(* IEC 61131-3 sources: Elmo_Master/Lasal_PRG/Elmo_EtherCAT_Test_4Axis/Network, 1 file *)

(* ---- ConfigObjects.st ---- *)
FUNCTION GLOBAL TAB TASK_CONF
_K_TASK, _K_REAL,
_K_END_VAR,

_K_TASK, _K_CYCLIC,
_K_END_VAR,

_K_TASK, _K_BACKGROUND,
_K_END_VAR,

_K_END_CONF
END_FUNCTION

FUNCTION GLOBAL TAB IPR_CONF
_K_IPR
	0$UINT,
_K_END_VAR,
_K_END_CONF
END_FUNCTION

FUNCTION GLOBAL TAB CONFIG_TABLES
00121$UINT,
0$UINT, 1, 58, "_AXISBASE",
0$UINT, 0, 5, "_CAN",
0$UINT, 1, 11, "_CANLIB",
0$UINT, 1, 0, "_CHECKSUM",
0$UINT, 1, 20, "_FILESYS",
0$UINT, 0, 5, "_LINKER",
0$UINT, 1, 0, "_LMCABSENCODER",
0$UINT, 1, 120, "_LMCAXIS",
0$UINT, 2, 111, "_LMCAXISBASE",
0$UINT, 1, 32, "_LMCAXISREF",
0$UINT, 1, 42, "_LMCAXISVIS",
0$UINT, 1, 63, "_LMCAXISVISINT",
0$UINT, 1, 0, "_LMCAXISVISLOGHANDLE",
0$UINT, 1, 0, "_LMCAXISVISLOGVIEWER",
0$UINT, 1, 13, "_LMCAXISVISPARA",
0$UINT, 1, 2, "_LMCAXISVOVMONITORING",
0$UINT, 1, 18, "_LMCBASECOORD",
0$UINT, 1, 7, "_LMCBELTAXIS",
0$UINT, 1, 5, "_LMCCALCMODELBASE",
0$UINT, 1, 2, "_LMCCALCMODELCONTROLLER",
0$UINT, 1, 24, "_LMCMATH_SO3",
0$UINT, 1, 75, "_LMCMATHFUNCTIONS",
0$UINT, 1, 1, "_LMCMODULEBASE",
0$UINT, 3, 0, "_LMCPROFILE",
0$UINT, 4, 0, "_LMCPROFILEBASE",
0$UINT, 1, 53, "_LMCPROFILEBUFFER",
0$UINT, 1, 44, "_LMCPROFILELOG",
0$UINT, 1, 30, "_LMCPROFILEVIS",
0$UINT, 1, 20, "_LMCPROFILEVISAXIS",
0$UINT, 1, 41, "_LMCPROFILEVISINT",
0$UINT, 1, 30, "_LMCPROFILEVISMOVEPARA",
0$UINT, 1, 0, "_LMCPUBLISHER",
0$UINT, 1, 11, "_LMCREFBASE",
0$UINT, 2, 22, "_LMCROBOTBASE",
0$UINT, 1, 42, "_LMCROBOTLOG",
0$UINT, 1, 21, "_LMCSAFETY",
0$UINT, 1, 2, "_LMCSPLINEBUFFER",
0$UINT, 1, 23, "_LMCTABLEBUFFER",
0$UINT, 1, 3, "_LMCTOOL",
0$UINT, 1, 1, "_MULTITASK",
0$UINT, 0, 5, "_OSKERNEL",
0$UINT, 1, 36, "_SERLIB",
0$UINT, 2, 0, "_STDLIB",
0$UINT, 1, 4, "_SYNCMEASURE",
0$UINT, 1, 3, "_SYNCMEASUREECAT",
0$UINT, 1, 1, "_TASKOBJECTCONTROL",
0$UINT, 1, 2, "_TCPIPSERVER",
0$UINT, 1, 1, "_TCPIPSERVERINTERFACE",
0$UINT, 1, 2, "_UDPTRANSCEIVER",
0$UINT, 1, 3, "_UDPTRANSCEIVERINTERFACE",
0$UINT, 1, 21, "ASCII_BIN",
0$UINT, 2, 2, "BUSINTERFACESDIASINTERNAL",
0$UINT, 1, 47, "CONTROLLER",
0$UINT, 1, 1, "CP313_IOS",
0$UINT, 1, 0, "CP733_IOS",
0$UINT, 0, 4, "CRITICALSECTION",
0$UINT, 2, 34, "DIASMASTER",
0$UINT, 1, 84, "DIASMASTERC",
0$UINT, 2, 26, "DIASMASTERMAIN",
0$UINT, 1, 1, "DIASMASTERPOSTSCAN",
0$UINT, 1, 2, "ECAT_DS402BASE",
0$UINT, 2, 3, "ECAT_MASTER_BASE",
0$UINT, 2, 1, "ECAT_SLAVE_BASE",
0$UINT, 1, 1, "ECAT_SLOTBASE",
0$UINT, 1, 2, "ECAT_SLOTMNG",
0$UINT, 1, 12, "EEPROM",
0$UINT, 0, 0, "ELMO_1",
0$UINT, 0, 0, "ELMO_2",
0$UINT, 0, 0, "ELMO_3",
0$UINT, 0, 0, "ELMO_4",
0$UINT, 1, 2, "ETHERCAT_HUB_BASE",
0$UINT, 2, 2, "ETHERCAT_PLC",
0$UINT, 1, 1, "ETHERCAT_SDOBASE",
0$UINT, 1, 1, "ETHERCATSLOT_HUB_BASE",
0$UINT, 1, 5, "GETCILINTERFACE",
0$UINT, 0, 0, "GL_9086_1",
0$UINT, 0, 0, "GL_9086_1_SLOT00",
0$UINT, 0, 0, "GL_9086_1_SLOT01",
0$UINT, 1, 22, "HUB_BASE",
0$UINT, 2, 12, "HUB_BASE_ROOT",
0$UINT, 2, 37, "HWBASE",
0$UINT, 2, 57, "HWBASECDIAS",
0$UINT, 1, 1, "HWCLOGGING",
0$UINT, 6, 0, "HWCONTROL",
0$UINT, 1, 11, "HWCONTROLBASE",
0$UINT, 1, 1, "HWRTPOSTSCAN",
0$UINT, 1, 7, "I2CCDIAS",
0$UINT, 0, 0, "LMCCONTROLCOMMANDSERVICE",
0$UINT, 0, 0, "LMCDIAGNOSTICSSERVICE",
0$UINT, 0, 0, "LMCECATINPUTLATCH",
0$UINT, 0, 0, "LMCRECORDERSTORE",
0$UINT, 0, 0, "LMCSDOEXECUTOR",
0$UINT, 0, 0, "LMCSETPOSITIONSTORE",
0$UINT, 0, 0, "LMCUDPCALLBACKSENDER",
0$UINT, 1, 0, "MERKER",
0$UINT, 1, 22, "MERKEREX",
0$UINT, 1, 0, "MOVESPLINETABLE",
0$UINT, 2, 77, "POSCONTROLLER",
0$UINT, 1, 9, "RAMFILE",
0$UINT, 3, 20, "SAFETYCDIAS_BASE",
0$UINT, 3, 0, "SAFETYMANAGER",
0$UINT, 1, 0, "SAFETYROUTINGTABLES",
0$UINT, 1, 5, "SAFETYUDP",
0$UINT, 2, 0, "SDIASBASE",
0$UINT, 1, 11, "SDIASHUBBASE",
0$UINT, 1, 100, "SDIASMANAGER",
0$UINT, 2, 8, "SDIASPLC",
0$UINT, 0, 46, "SIGCLIB",
0$UINT, 1, 11, "STRING",
0$UINT, 1, 86, "STRINGINTERNAL",
0$UINT, 1, 22, "SYNCCALL",
0$UINT, 0, 0, "TCPIPSERVER",
0$UINT, 0, 0, "TCPMOTIONINTERFACE",
0$UINT, 2, 22, "VARAN_BASE",
0$UINT, 3, 9, "VARANMANAGER",
0$UINT, 2, 8, "VARANMANAGER_1",
0$UINT, 2, 10, "VARANMANAGER_2",
0$UINT, 1, 27, "VARANMANAGER_BASE",
0$UINT, 1, 3, "VIRTUALBASEINIT",
0$UINT, 2, 12, "WATCHDOGDIAS",
0$UINT, 1, 4, "XXXBASE_IOS",
ONE_CFG$UINT, 0, 0, "ONE_Comm_Network",
ONE_CFG$UINT, 0, 0, "ONE_EtherCAT_Network",
ONE_CFG$UINT, 0, 0, "ONE_HW_Network",
ONE_CFG$UINT, 0, 0, "ONE_Motion_Network",
TASK_CFG$UINT, 0, 0, "TASK_CONF",
IPR_CFG$UINT, 0, 0, "IPR_CONF",
PRJ_CFG$UINT, 0, 0, "Elmo_EtherCAT_Test_4Axis",
END_FUNCTION

#ifdef __LSLLDR_IOELEMENTS__
FUNCTION GLOBAL TAB _IO_ELEMENTS_TAB
0001$UINT, 0001$UINT,
"**IOCONN_EMPTY**", "Elmo_11.AxError",
0044$UINT,
"**IOCONN_EMPTY**", "PosController1.iHWErrors",
"**IOCONN_EMPTY**", "PosController1.HWErrorQuit",
"**IOCONN_EMPTY**", "PosController1.oActive",
"**IOCONN_EMPTY**", "PosController1.oOutputSignal",
"**IOCONN_EMPTY**", "PosController1.DriveEnabled",
"**IOCONN_EMPTY**", "_LMCAxis1.ActPosition",
"**IOCONN_EMPTY**", "_LMCAxis1.HWError",
"**IOCONN_EMPTY**", "_LMCAxis1.HWReady",
"**IOCONN_EMPTY**", "PosController2.iHWErrors",
"**IOCONN_EMPTY**", "PosController2.HWErrorQuit",
"**IOCONN_EMPTY**", "PosController2.oActive",
"**IOCONN_EMPTY**", "PosController2.oOutputSignal",
"**IOCONN_EMPTY**", "PosController2.DriveEnabled",
"**IOCONN_EMPTY**", "_LMCAxis2.ActPosition",
"**IOCONN_EMPTY**", "_LMCAxis2.HWError",
"**IOCONN_EMPTY**", "_LMCAxis2.HWReady",
"**IOCONN_EMPTY**", "PosController3.iHWErrors",
"**IOCONN_EMPTY**", "PosController3.HWErrorQuit",
"**IOCONN_EMPTY**", "PosController3.oActive",
"**IOCONN_EMPTY**", "PosController3.oOutputSignal",
"**IOCONN_EMPTY**", "PosController3.DriveEnabled",
"**IOCONN_EMPTY**", "_LMCAxis3.ActPosition",
"**IOCONN_EMPTY**", "_LMCAxis3.HWError",
"**IOCONN_EMPTY**", "_LMCAxis3.HWReady",
"**IOCONN_EMPTY**", "PosController4.iHWErrors",
"**IOCONN_EMPTY**", "PosController4.HWErrorQuit",
"**IOCONN_EMPTY**", "PosController4.oActive",
"**IOCONN_EMPTY**", "PosController4.oOutputSignal",
"**IOCONN_EMPTY**", "PosController4.DriveEnabled",
"**IOCONN_EMPTY**", "_LMCAxis4.ActPosition",
"**IOCONN_EMPTY**", "_LMCAxis4.HWError",
"**IOCONN_EMPTY**", "_LMCAxis4.HWReady",
"**IOCONN_EMPTY**", "LMCEcatInputLatch1.EcatMaster",
"**IOCONN_EMPTY**", "LMCEcatInputLatch1.Drive1",
"**IOCONN_EMPTY**", "LMCEcatInputLatch1.Drive2",
"**IOCONN_EMPTY**", "LMCEcatInputLatch1.Drive3",
"**IOCONN_EMPTY**", "LMCEcatInputLatch1.Drive4",
"**IOCONN_EMPTY**", "LMCSdoExecutor1.toSlave",
"**IOCONN_EMPTY**", "LMCEcatInputLatch1.Coupler",
"**IOCONN_EMPTY**", "LMCEcatInputLatch1.InputSlot",
"**IOCONN_EMPTY**", "LMCEcatInputLatch1.OutputSlot",
"**IOCONN_EMPTY**", "LMCSdoExecutor2.toSlave",
"**IOCONN_EMPTY**", "LMCSdoExecutor3.toSlave",
"**IOCONN_EMPTY**", "LMCSdoExecutor4.toSlave",
END_FUNCTION
#endif //__LSLLDR_IOELEMENTS__

FUNCTION GLOBAL TAB CH_REDIRECT_EMB_TAB
0000$UINT,
00030$UINT,
"_TCPIPSERVER;SEMANAME01", "\STRSEMANAME01.DATA",
"_TCPIPSERVER;SEMANAME02", "\STRSEMANAME02.DATA",
"_TCPIPSERVER;TASKNAME", "\STRTASKNAME.DATA",
"ECAT_DS402BASE;DEVICENAME", "\DEVICENAMESTR.DATA",
"ECAT_DS402BASE;PRODUCTREVISION", "\PRODUCTREVSTR.DATA",
"ECAT_MASTER_BASE;SOFTWAREVERSION", "\STRSOFTWAREVERSION.DATA",
"ECAT_SLAVE_BASE;DEVICENAME", "\DEVICENAMESTR.DATA",
"ECAT_SLAVE_BASE;PRODUCTREVISION", "\PRODUCTREVSTR.DATA",
"ECAT_SLOTMNG;DEVICENAME", "\DEVICENAMESTR.DATA",
"ECAT_SLOTMNG;PRODUCTREVISION", "\PRODUCTREVSTR.DATA",
"ELMO_1;DEVICENAME", "\DEVICENAMESTR.DATA",
"ELMO_1;PRODUCTREVISION", "\PRODUCTREVSTR.DATA",
"ELMO_2;DEVICENAME", "\DEVICENAMESTR.DATA",
"ELMO_2;PRODUCTREVISION", "\PRODUCTREVSTR.DATA",
"ELMO_3;DEVICENAME", "\DEVICENAMESTR.DATA",
"ELMO_3;PRODUCTREVISION", "\PRODUCTREVSTR.DATA",
"ELMO_4;DEVICENAME", "\DEVICENAMESTR.DATA",
"ELMO_4;PRODUCTREVISION", "\PRODUCTREVSTR.DATA",
"ETHERCAT_PLC;SOFTWAREVERSION", "\STRSOFTWAREVERSION.DATA",
"ETHERCAT_SDOBASE;PARASTRING", "\STRSDOPARASTRING.DATA",
"GL_9086_1;DEVICENAME", "\DEVICENAMESTR.DATA",
"GL_9086_1;PRODUCTREVISION", "\PRODUCTREVSTR.DATA",
"HWBASECDIAS;SERIALNO", "\SERIALNOSTR.DATA",
"LMCSDOEXECUTOR;PARASTRING", "\STRSDOPARASTRING.DATA",
"SAFETYCDIAS_BASE;SERIALNO", "\SERIALNOSTR.DATA",
"SDIASBASE;SERIALNO", "\SERIALNOSTR.DATA",
"TCPIPSERVER;SEMANAME01", "\STRSEMANAME01.DATA",
"TCPIPSERVER;SEMANAME02", "\STRSEMANAME02.DATA",
"TCPIPSERVER;TASKNAME", "\STRTASKNAME.DATA",
"VARAN_BASE;SERIALNO", "\SERIALNOSTR.DATA",
END_FUNCTION
